// TIA Portal V21 export
// export: Created 2026-11-11T00:47:53.6687691Z, ExportSetting WithDefaults, DisplayName Totally Integrated Automation Portal, DisplayVersion V21 Update 3, DisplayName STEP 7 Professional, DisplayVersion V21 Update 3, DisplayName STEP 7 Safety, DisplayVersion V21, DisplayName Tech WebApplication, DisplayVersion V21, DisplayName WinCC Basic/Comfort/Advanced, DisplayVersion V21 Update 3, DisplayName WinCC Unified, DisplayVersion V21 Update 3
FUNCTION_BLOCK "FB_Lad_ex059"   // FB396, LAD
{ S7_Optimized_Access := 'TRUE' }
VERSION : 0.1
// stored: AutoNumber true, IsIECCheckEnabled false, IsRetainMemResEnabled false, MemoryReserve 100, SetENOAutomatically false, UDAEnableTagReadback false
   VAR_INPUT
      v_req : Bool;
      v_laddr : HW_IO;
      v_recnum : Byte;
      v_record : Variant;
   END_VAR
   VAR_OUTPUT
      v_ret_val : Int;
      v_busy : Bool;
   END_VAR
BEGIN

REGION Network 1: WR_REC - Write data record to I/O
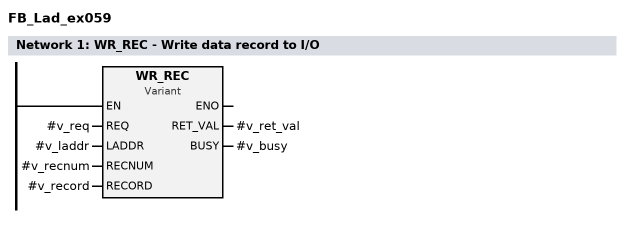
   RUNG wire#powerrail
      { S7_Templates := "[card := 0, ptr_type := Variant, laddr_type := HW_IO]" } WR_REC(REQ := #v_req, LADDR := #v_laddr, RECNUM := #v_recnum, RECORD := #v_record, RET_VAL => #v_ret_val, BUSY => #v_busy)
   END_RUNG
   // the same network as SCL:
   #v_ret_val := WR_REC(REQ := #v_req,
                        LADDR := #v_laddr,
                        RECNUM := #v_recnum,
                        RECORD := #v_record,
                        BUSY => #v_busy);
END_REGION
END_FUNCTION_BLOCK
